(* CODESYS project StyleProbe.export

Project tree, tasks and I/O mapping:
  visualisation StyleProbe
*)

// /StyleProbe
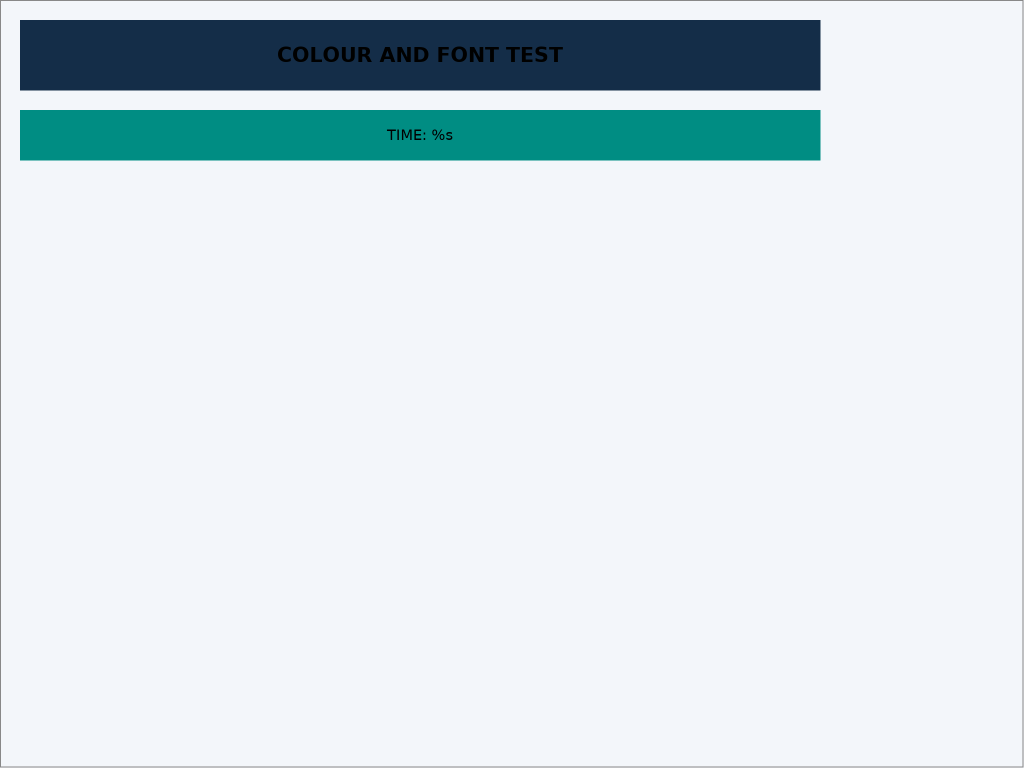
VISUALIZATION StyleProbe  // 1024x768
    Rectangle (0,0 1024x768)
    Rectangle (20,20 800x70), "COLOUR AND FONT TEST"
    Rectangle (20,110 800x50), "TIME: %s", text variable: Team_HMI.sDateTime
END_VISUALIZATION
